Fanuc KAREL source: KO00001.KL

PROGRAM KO00001
%NOLOCKGROUP
VAR
  P1: POSITION
  P2: POSITION
  P3: POSITION
  OUT: POSITION
BEGIN
  OUT = FRAME(P1, P2, P3)
END KO00001
